Fanuc KAREL source: kt00071.KL

-- PROVISIONAL review KL for V940-1; original PC SHA256 34aa6e6533cbc01e1f37b9fb42413d47a8d10e5cf0a362d3acce451b8b4f4d49
-- Incomplete behavior may be omitted. Consult companion uncertainty JSON. Do not deploy.
PROGRAM KT00071
%NOLOCKGROUP
VAR
  I1 : INTEGER
  OUT : INTEGER
-- UNRESOLVED_DECL H2 type=002017
BEGIN
  -- V9_ZERO_TABLE_METADATA_HINT layout=0001; no indexed target words; source/name/runtime held
  -- UNRESOLVED_PC offsets 5-16; opcodes 2E,23
  -- UNRESOLVED_PC offsets 21-35; opcodes 2E,22,9D,33,B4
  -- UNRESOLVED_PC offsets 40-62; opcodes 21,22,9D,33,B3,54,23
  -- UNRESOLVED_PC offsets 67-71; opcodes 7F
END KT00071
